TYPE TYPE_SEQUENCE :
STRUCT
	active : BOOL;
	lineNo : UDINT;
	task : ARRAY[0..Size.MAX_TASK-1] OF TYPE_TASK;
END_STRUCT
END_TYPE

(* stored: Version 1.1.0.1, ProductVersion 3.1.4024.12
   DUT TYPE_SEQUENCE: Id {68362961-54be-48b5-b292-de01a2e92ee2} *)
